{region 'Documentation'}
(*!
<summary>Checks REAL absolute tolerance boundaries and Error escalation in both relations.</summary>
<description>
Named rows separate independent comparisons by a disabled reset call.
Only explicitly marked escalation rows retain the preceding subject result.
Outer Assertions latch every observation before advancing to the next row.
All finite comparison values are exact binary fractions; expected results are literal.
ErrorAfterEqualFailure and ErrorAfterNotEqualFailure exercise each held-Failed guard.
RepeatedError and ValidInputsAfterError require held Error without another finding.
Intentional findings remain in the local capture; no production algorithm is copied.
</description>
*)
{endregion}
FUNCTION_BLOCK Test_AssertionTolerance_Real EXTENDS TestCaseBase
VAR
    FEqualSubject : AssertEqualTolerance_Real;
    FNotEqualSubject : AssertNotEqualTolerance_Real;
    FActual : REAL;
    FExpected : REAL;
    FTolerance : REAL;
    FExpectedEqualResult : E_Result;
    FExpectedNotEqualResult : E_Result;
    FExpectedFindings : UDINT;
    FExpectedEqualFinding : E_Result;
    FExpectedNotEqualFinding : E_Result;
    FCapture : EventBuffer;
    FEvents : ARRAY[1..CaptureLength] OF ST_Event;
    FCaptureFifo : ST_FifoStatus;
    FCaptureStatus : ST_EventBufferStatus;
    FRow : UINT;
    FRowPrepared : BOOL;
    FPreserveResults : BOOL;
    FObservationReady : BOOL;
    FChecked : BOOL;
    FSetupValid : BOOL;
END_VAR
VAR
    FEqualResult : AssertTrue;
    FEqualResultMatches : BOOL;
    FNotEqualResult : AssertTrue;
    FNotEqualResultMatches : BOOL;
    FCaptureIntegrity : AssertTrue;
    FCaptureIntegrityMatches : BOOL;
    FFindingDetails : AssertTrue;
    FFindingDetailsMatch : BOOL;
END_VAR
VAR CONSTANT
    CaptureLength : UINT := 8;
    EqualValues : UINT := 1;
    InsideLower : UINT := 2;
    InsideUpper : UINT := 3;
    AtLowerBoundary : UINT := 4;
    AtUpperBoundary : UINT := 5;
    OutsideLower : UINT := 6;
    OutsideUpper : UINT := 7;
    ZeroToleranceEqual : UINT := 8;
    ZeroToleranceDifferent : UINT := 9;
    NegativeTolerance : UINT := 10;
    EqualFailureBeforeError : UINT := 11;
    ErrorAfterEqualFailure : UINT := 12;
    RepeatedError : UINT := 13;
    ValidInputsAfterError : UINT := 14;
    NotEqualFailureBeforeError : UINT := 15;
    ErrorAfterNotEqualFailure : UINT := 16;
    ResetRestoresEvaluation : UINT := 17;
    LastRow : UINT := ResetRestoresEvaluation;
END_VAR

SUPER^();

{region 'Documentation'}
(*!
<summary>Collects only outer checking Assertions, never intentional subject findings.</summary>
*)
{endregion}
METHOD PROTECTED AggregateResults
VAR_INPUT
    Aggregator : I_ResultAggregator; //! Borrowed result sink owned by the outer Test Case; add this test's checking Assertions without resetting or retaining the sink.
END_VAR
Aggregator.AddProvider(Provider := FEqualResult);
Aggregator.AddProvider(Provider := FNotEqualResult);
Aggregator.AddProvider(Provider := FCaptureIntegrity);
Aggregator.AddProvider(Provider := FFindingDetails);
END_METHOD

{region 'Documentation'}
(*!
<summary>Calls each inherited production Assertion once using the selected row.</summary>
*)
{endregion}
METHOD PRIVATE CallSubjects
VAR_INPUT
    Enable : BOOL; //! Observation-enable input forwarded to the controlled Assertion subjects for this call.
END_VAR
FEqualSubject(Enable := Enable,
    State := E_State.Running,
    IN := FActual,
    Expected := FExpected,
    Tolerance := FTolerance);
FNotEqualSubject(Enable := Enable,
    State := E_State.Running,
    IN := FActual,
    Expected := FExpected,
    Tolerance := FTolerance);
END_METHOD

{region 'Documentation'}
(*!
<summary>Extends base validation with subject and checking-Assertion setup.</summary>
*)
{endregion}
METHOD PROTECTED CheckInitialization : BOOL //! TRUE when the inherited initialization check and this concrete fixture check both accept the setup.
CheckInitialization := SUPER^.CheckInitialization();
IF NOT CheckInitialization THEN
    RETURN;
END_IF;

CheckInitialization := FSetupValid
    AND FEqualResult.IsInitialized
    AND FNotEqualResult.IsInitialized
    AND FCaptureIntegrity.IsInitialized
    AND FFindingDetails.IsInitialized;
IF NOT CheckInitialization THEN
    EventPublisher.PublishEvent(Event := CreateFrameworkEvent(Name := Name,
        ResourceName := '',
        State := State,
        Severity := E_EventSeverity.Error,
        Message := 'Tolerance selftest setup failed.'));
END_IF;
END_METHOD

{region 'Documentation'}
(*!
<summary>Checks literal results, finding count and isolated finding identities.</summary>
*)
{endregion}
METHOD PRIVATE CheckResults
VAR
    FindingIndex : UINT;
    NotEqualFindingMatches : BOOL;
END_VAR
FEqualResultMatches := FEqualSubject.Result = FExpectedEqualResult;
FNotEqualResultMatches := FNotEqualSubject.Result = FExpectedNotEqualResult;
FCaptureIntegrityMatches := (FCaptureStatus.SequenceId = FExpectedFindings)
    AND (FCaptureStatus.LostEventCount = 0);

FindingIndex := 1;
FFindingDetailsMatch := TRUE;
IF FExpectedEqualFinding <> E_Result.NotEvaluated THEN
    FFindingDetailsMatch := IsFindingValid(Index := FindingIndex,
        ExpectedName := FEqualSubject.Name,
        ExpectedResult := FExpectedEqualFinding);
    FindingIndex := FindingIndex + 1;
END_IF;
IF FExpectedNotEqualFinding <> E_Result.NotEvaluated THEN
    NotEqualFindingMatches := IsFindingValid(Index := FindingIndex,
        ExpectedName := FNotEqualSubject.Name,
        ExpectedResult := FExpectedNotEqualFinding);
    FFindingDetailsMatch := FFindingDetailsMatch AND NotEqualFindingMatches;
END_IF;
END_METHOD

{region 'Documentation'}
(*!
<summary>Configures checking Assertions; subject actions remain in the test script.</summary>
*)
{endregion}
METHOD PROTECTED Configure
VAR
    Initialized : BOOL;
END_VAR
FPreparationStateCount := 0;
FTestStateCount := 1;
FEqualResult.Initialize(Parent := THIS^,
    AssertionName := 'EqualResult');
FNotEqualResult.Initialize(Parent := THIS^,
    AssertionName := 'NotEqualResult');
FCaptureIntegrity.Initialize(Parent := THIS^,
    AssertionName := 'CaptureIntegrity');
FFindingDetails.Initialize(Parent := THIS^,
    AssertionName := 'FindingDetails');
FSetupValid := FCapture.Initialize(Buffer := FEvents,
    FifoControl := FCaptureFifo,
    Status := FCaptureStatus);
FEqualSubject.BindPublisher(Publisher := FCapture);
Initialized := FEqualSubject.Initialize(Parent := THIS^,
    AssertionName := 'EqualSubject');
FSetupValid := FSetupValid AND Initialized;
FNotEqualSubject.BindPublisher(Publisher := FCapture);
Initialized := FNotEqualSubject.Initialize(Parent := THIS^,
    AssertionName := 'NotEqualSubject');
FSetupValid := FSetupValid AND Initialized;
END_METHOD

{region 'Documentation'}
(*!
<summary>Reads one of at most two captured findings; caller supplies index 1 or 2.</summary>
*)
{endregion}
METHOD PRIVATE IsFindingValid : BOOL //! TRUE when the selected captured finding satisfies the scenario metadata and diagnostic checks.
VAR_INPUT
    Index : UINT; //! One-based index in the retained isolated event capture.
    ExpectedName : STRING(GVL_Constants.NameLength); //! Independently authored Assertion name expected in the selected finding.
    ExpectedResult : E_Result; //! Independently authored finding result.
END_VAR
IsFindingValid := (FEvents[Index].SequenceId = UINT_TO_UDINT(Index))
    AND (FEvents[Index].Name = ExpectedName)
    AND (FEvents[Index].OwnerScope = E_OwnerScope.Assertion)
    AND (FEvents[Index].EventType = E_EventType.Result)
    AND (FEvents[Index].State = E_State.Running)
    AND (FEvents[Index].Result = ExpectedResult)
    AND (FEvents[Index].Message <> '');
END_METHOD

{region 'Documentation'}
(*!
<summary>Completes abort without asynchronous resources.</summary>
*)
{endregion}
METHOD PROTECTED ProcessAbort
VAR_INPUT
    Enable : BOOL; //! Phase permission supplied by the owning Test Case; FALSE does not authorize progression, while observation may continue.
END_VAR
IF Enable THEN
    CompleteAbort();
END_IF;
END_METHOD

{region 'Documentation'}
(*!
<summary>Latches checked observations before the next script step may proceed.</summary>
*)
{endregion}
METHOD PROTECTED ProcessAssertions
VAR_INPUT
    Enable : BOOL; //! Phase permission supplied by the owning Test Case; FALSE does not authorize progression, while observation may continue.
END_VAR
VAR
    Evaluate : BOOL;
END_VAR
Evaluate := Enable AND FObservationReady;
FEqualResult(Enable := Evaluate,
    State := State,
    IN := FEqualResultMatches);
FNotEqualResult(Enable := Evaluate,
    State := State,
    IN := FNotEqualResultMatches);
FCaptureIntegrity(Enable := Evaluate,
    State := State,
    IN := FCaptureIntegrityMatches);
FFindingDetails(Enable := Evaluate,
    State := State,
    IN := FFindingDetailsMatch);
IF Evaluate THEN
    FChecked := TRUE;
END_IF;
END_METHOD

{region 'Documentation'}
(*!
<summary>No Preparation phase is required.</summary>
*)
{endregion}
METHOD PROTECTED ProcessPreparations
VAR_INPUT
    // SA0033: Required hook; this test has no Preparation phase.
    {attribute 'analysis' := '-33'}
    Enable : BOOL; //! Phase permission supplied by the owning Test Case; FALSE does not authorize progression, while observation may continue.
END_VAR
END_METHOD

{region 'Documentation'}
(*!
<summary>Restarts the script and resets the checking Assertions.</summary>
*)
{endregion}
METHOD PROTECTED ProcessReset
FRow := EqualValues;
FRowPrepared := FALSE;
FChecked := FALSE;
FObservationReady := FALSE;
FEqualResult.Reset();
FEqualResultMatches := TRUE;
FNotEqualResult.Reset();
FNotEqualResultMatches := TRUE;
FCaptureIntegrity.Reset();
FCaptureIntegrityMatches := TRUE;
FFindingDetails.Reset();
FFindingDetailsMatch := TRUE;
CompleteReset();
END_METHOD

{region 'Documentation'}
(*!
<summary>Advances one bounded script step per active PLC cycle.</summary>
*)
{endregion}
METHOD PROTECTED ProcessTests
VAR_INPUT
    Enable : BOOL; //! Phase permission supplied by the owning Test Case; FALSE does not authorize progression, while observation may continue.
END_VAR
IF NOT Enable THEN
    RETURN;
END_IF;

IF FChecked THEN
    FChecked := FALSE;
    FObservationReady := FALSE;
    IF FRow = LastRow THEN
        CompleteTests();
        RETURN;
    END_IF;
    FRow := FRow + 1;
    FRowPrepared := FALSE;
END_IF;

IF NOT FRowPrepared THEN
    SelectRow();
    FCapture.Reset();
    IF NOT FPreserveResults THEN
        ResetSubjects();
    END_IF;
    CallSubjects(Enable := FALSE);
    FRowPrepared := TRUE;
ELSE
    CallSubjects(Enable := TRUE);
    CheckResults();
    FObservationReady := TRUE;
END_IF;
END_METHOD

{region 'Documentation'}
(*!
<summary>Requests fresh subject results before the next disabled call.</summary>
*)
{endregion}
METHOD PRIVATE ResetSubjects
FEqualSubject.Reset();
FNotEqualSubject.Reset();
END_METHOD

{region 'Documentation'}
(*!
<summary>Selects literal expectations; only named escalation rows retain preceding subject results.</summary>
*)
{endregion}
METHOD PRIVATE SelectRow
FPreserveResults := FALSE;
FExpected := REAL#8.0;
CASE FRow OF
    EqualValues:
        FActual := REAL#8.0;
        FTolerance := REAL#0.5;
        FExpectedEqualResult := E_Result.Passed;
        FExpectedNotEqualResult := E_Result.Failed;
        FExpectedFindings := 1;
        FExpectedEqualFinding := E_Result.NotEvaluated;
        FExpectedNotEqualFinding := E_Result.Failed;
    InsideLower:
        FActual := REAL#7.75;
        FTolerance := REAL#0.5;
        FExpectedEqualResult := E_Result.Passed;
        FExpectedNotEqualResult := E_Result.Failed;
        FExpectedFindings := 1;
        FExpectedEqualFinding := E_Result.NotEvaluated;
        FExpectedNotEqualFinding := E_Result.Failed;
    InsideUpper:
        FActual := REAL#8.25;
        FTolerance := REAL#0.5;
        FExpectedEqualResult := E_Result.Passed;
        FExpectedNotEqualResult := E_Result.Failed;
        FExpectedFindings := 1;
        FExpectedEqualFinding := E_Result.NotEvaluated;
        FExpectedNotEqualFinding := E_Result.Failed;
    AtLowerBoundary:
        FActual := REAL#7.5;
        FTolerance := REAL#0.5;
        FExpectedEqualResult := E_Result.Passed;
        FExpectedNotEqualResult := E_Result.Failed;
        FExpectedFindings := 1;
        FExpectedEqualFinding := E_Result.NotEvaluated;
        FExpectedNotEqualFinding := E_Result.Failed;
    AtUpperBoundary:
        FActual := REAL#8.5;
        FTolerance := REAL#0.5;
        FExpectedEqualResult := E_Result.Passed;
        FExpectedNotEqualResult := E_Result.Failed;
        FExpectedFindings := 1;
        FExpectedEqualFinding := E_Result.NotEvaluated;
        FExpectedNotEqualFinding := E_Result.Failed;
    OutsideLower:
        FActual := REAL#7.25;
        FTolerance := REAL#0.5;
        FExpectedEqualResult := E_Result.Failed;
        FExpectedNotEqualResult := E_Result.Passed;
        FExpectedFindings := 1;
        FExpectedEqualFinding := E_Result.Failed;
        FExpectedNotEqualFinding := E_Result.NotEvaluated;
    OutsideUpper:
        FActual := REAL#8.75;
        FTolerance := REAL#0.5;
        FExpectedEqualResult := E_Result.Failed;
        FExpectedNotEqualResult := E_Result.Passed;
        FExpectedFindings := 1;
        FExpectedEqualFinding := E_Result.Failed;
        FExpectedNotEqualFinding := E_Result.NotEvaluated;
    ZeroToleranceEqual:
        FActual := REAL#8.0;
        FTolerance := REAL#0.0;
        FExpectedEqualResult := E_Result.Passed;
        FExpectedNotEqualResult := E_Result.Failed;
        FExpectedFindings := 1;
        FExpectedEqualFinding := E_Result.NotEvaluated;
        FExpectedNotEqualFinding := E_Result.Failed;
    ZeroToleranceDifferent:
        FActual := REAL#8.25;
        FTolerance := REAL#0.0;
        FExpectedEqualResult := E_Result.Failed;
        FExpectedNotEqualResult := E_Result.Passed;
        FExpectedFindings := 1;
        FExpectedEqualFinding := E_Result.Failed;
        FExpectedNotEqualFinding := E_Result.NotEvaluated;
    NegativeTolerance:
        FActual := REAL#8.0;
        FTolerance := REAL#-0.5;
        FExpectedEqualResult := E_Result.Error;
        FExpectedNotEqualResult := E_Result.Error;
        FExpectedFindings := 2;
        FExpectedEqualFinding := E_Result.Error;
        FExpectedNotEqualFinding := E_Result.Error;
    EqualFailureBeforeError:
        FActual := REAL#9.0;
        FTolerance := REAL#0.5;
        FExpectedEqualResult := E_Result.Failed;
        FExpectedNotEqualResult := E_Result.Passed;
        FExpectedFindings := 1;
        FExpectedEqualFinding := E_Result.Failed;
        FExpectedNotEqualFinding := E_Result.NotEvaluated;
    ErrorAfterEqualFailure:
        FActual := REAL#9.0;
        FTolerance := REAL#-0.5;
        FExpectedEqualResult := E_Result.Error;
        FExpectedNotEqualResult := E_Result.Error;
        FExpectedFindings := 2;
        FExpectedEqualFinding := E_Result.Error;
        FExpectedNotEqualFinding := E_Result.Error;
        FPreserveResults := TRUE;
    RepeatedError:
        FActual := REAL#9.0;
        FTolerance := REAL#-0.5;
        FExpectedEqualResult := E_Result.Error;
        FExpectedNotEqualResult := E_Result.Error;
        FExpectedFindings := 0;
        FExpectedEqualFinding := E_Result.NotEvaluated;
        FExpectedNotEqualFinding := E_Result.NotEvaluated;
        FPreserveResults := TRUE;
    ValidInputsAfterError:
        FActual := REAL#8.0;
        FTolerance := REAL#0.5;
        FExpectedEqualResult := E_Result.Error;
        FExpectedNotEqualResult := E_Result.Error;
        FExpectedFindings := 0;
        FExpectedEqualFinding := E_Result.NotEvaluated;
        FExpectedNotEqualFinding := E_Result.NotEvaluated;
        FPreserveResults := TRUE;
    NotEqualFailureBeforeError:
        FActual := REAL#8.0;
        FTolerance := REAL#0.5;
        FExpectedEqualResult := E_Result.Passed;
        FExpectedNotEqualResult := E_Result.Failed;
        FExpectedFindings := 1;
        FExpectedEqualFinding := E_Result.NotEvaluated;
        FExpectedNotEqualFinding := E_Result.Failed;
    ErrorAfterNotEqualFailure:
        FActual := REAL#8.0;
        FTolerance := REAL#-0.5;
        FExpectedEqualResult := E_Result.Error;
        FExpectedNotEqualResult := E_Result.Error;
        FExpectedFindings := 2;
        FExpectedEqualFinding := E_Result.Error;
        FExpectedNotEqualFinding := E_Result.Error;
        FPreserveResults := TRUE;
    ResetRestoresEvaluation:
        FActual := REAL#8.0;
        FTolerance := REAL#0.5;
        FExpectedEqualResult := E_Result.Passed;
        FExpectedNotEqualResult := E_Result.Failed;
        FExpectedFindings := 1;
        FExpectedEqualFinding := E_Result.NotEvaluated;
        FExpectedNotEqualFinding := E_Result.Failed;
ELSE
    Error(Message := 'Unknown tolerance test row.');
END_CASE;
END_METHOD

END_FUNCTION_BLOCK

(* stored: Version 1.1.0.1
   POU Test_AssertionTolerance_Real: Id {b34d890e-c587-42a6-8634-10808ea1825f}, SpecialFunc None
   Folder Internal: Id {5dfa81a5-b51c-453c-8184-aef1b209c70f}
   Method AggregateResults: Id {58679063-c902-47b1-b330-b95450a2d106}
   Method CallSubjects: Id {1996fa2d-6714-4c60-bcf3-e0656991647d}
   Method CheckInitialization: Id {c60dd689-d452-4f79-b3ce-c87837609713}
   Method CheckResults: Id {5039f1b1-3d01-43b9-a1c1-858494927f3b}
   Method Configure: Id {f52535ea-9e9f-4c5f-93ba-c36d397788f4}
   Method IsFindingValid: Id {3e8e8bf2-9630-4fe2-89c4-a690b9224c68}
   Method ProcessAbort: Id {bda7e4bf-462b-4c6e-b048-7a2d966d48a4}
   Method ProcessAssertions: Id {baf3ea1d-41f4-402b-88fb-542fc86c22b2}
   Method ProcessPreparations: Id {a49a31cb-4380-4483-b7de-bc330ccbc0fe}
   Method ProcessReset: Id {66520a62-5326-454e-956e-d5ce285fc388}
   Method ProcessTests: Id {face6469-9197-4d6f-b281-aa02e3093142}
   Method ResetSubjects: Id {4b77ee09-386a-4ab0-9875-2517f1d1fec6}
   Method SelectRow: Id {908f3bca-701c-4a40-ab3d-0ab767922cb6} *)
